(* IEC 61131-3 sources: moqui-plc/simatic-ax/src/moqui/framework/src/main/org/moqui/context, 9 files *)

(* ---- LogCmd.st ---- *)
TYPE LogCmd : (
    Idle, (* Waiting for commands *)
    Push (* Inserting a new log entry *)
); END_TYPE

(* ---- LogEvent.st ---- *)
TYPE LogEvent : STRUCT
	(* Unique identifier for the log event *)
    logEventId : STRING;
    loggerName : STRING;
	marker : LogMarker;
    level : LogLevel;
    logEventDate : DATE_AND_TIME;
	source : STRING;
	payloadType : LogPayloadType;
    payload : LogPayload;
	(* contextData: STRING; *)
	(*
	 * Occurrences this record stands for: 1 for an event, N for the summary that LoggerFacade writes when the
	 * same event was repeated N more times inside the suppression window ("last message repeated N times").
	 *)
    repeatCount : UINT;
	(* Position of the record in its LogRingBuffer, set by the buffer: consecutive records of one source differ by 1. *)
	sequence : UDINT;
END_STRUCT; END_TYPE

(* ---- LogLevel.st ---- *)
TYPE LogLevel : (
	Trace,
	Debug,
	Info,
	Warn,
	Error,
	Fatal,
	All,
	Off
); END_TYPE

(* ---- LogMarker.st ---- *)
TYPE LogMarker : (
	Diagnostics,
	Lifecycle,
	Integration,
	Health,
	Telemetry,
	AuditLog,
	Kpi,
	Measurement
); END_TYPE

(* ---- LogPayload.st ---- *)
TYPE LogPayload : STRUCT
	message : STRING;
    enumValue : UINT;
    numericValue : LREAL;
END_STRUCT; END_TYPE

(* ---- LogPayloadType.st ---- *)
TYPE LogPayloadType : (
    Text,
	Numeric,
	Enum
); END_TYPE

(* ---- LogSource.st ---- *)
(*
 * One registered LoggerFacade buffer, as seen by its consumer.
 * LoggerFacade sets logRef once; every other field belongs to the consumer. The AX port has no MQTT consumer yet
 * (the intended Siemens path is OPC UA): a future consumer follows LogDispatcher of the canonical IEC source.
 *)
TYPE LogSource : STRUCT
	(* Reference to log ring buffer *)
    logRef : REF_TO LogRingBuffer;
	(* Slot of the oldest record not yet released by the consumer *)
	readSlot : UINT := UINT#1;
	(* LogRingBuffer.droppedCount already reported by the consumer *)
	reportedDropCount : UDINT;
	(* Records published, and records discarded by the consumer *)
	publishedCount : UDINT;
	discardedCount : UDINT;
END_STRUCT; END_TYPE

(* ---- LoggerFacade.st ---- *)
USING System.Strings;

(*
 * Logger with local circular buffer and duplicate suppression.
 * Designed for central orchestration by a global LogAppender.
 *
 * - Level threshold: events below the global logMinLevel are ignored, as a log4j logger level.
 * - Duplicate suppression: an event equal to the last stored one (same logger, source, level, marker, payload
 *   type and value) within suppressDuration is only counted. The count is written later as one summary record,
 *   a copy of the event with repeatCount = repetitions, when a different event arrives or when the window has
 *   elapsed at any later call ("last message repeated N times"). Stored records are never modified.
 * - Rate limit: at most maxEventsPerWindow new events are stored in one suppressDuration window. Further
 *   events are only counted; at the first call after the window one Warn event reports how many were suppressed.
 *   Repetitions counted by duplicate suppression do not count against the limit.
 * - The local LogRingBuffer has this block as its only producer: call it from one task only.
 * - Inputs are retained between calls, as for every function block: pass level at every call,
 *   otherwise the event gets the level of the previous call.
 * - Generated logEventId: loggerName-<event sequence> (AX: no millisecond clock is read for the ID).
 *)
FUNCTION_BLOCK LoggerFacade
	VAR_EXTERNAL CONSTANT
		defaultLogLevel : LogLevel;
		defaultLogSuppressDuration : TIME;
		defaultLogSuppressDuplicates : BOOL;
		defaultLogMaxEventsPerWindow : UINT;
		LOG_SOURCE_LIST_MAX_SIZE : UINT;
	END_VAR
	VAR_EXTERNAL
		logSourceList : ARRAY[1..LOG_SOURCE_LIST_MAX_SIZE] OF LogSource;
		logSourceListSize : DINT;
		logMinLevel : LogLevel;
	END_VAR
	(* Log event data *)
	VAR_INPUT
		enable : BOOL;
		logEventId : STRING := '';
		loggerName : STRING;
		level : LogLevel := defaultLogLevel;
		marker : LogMarker := LogMarker#Diagnostics;
		source : STRING;
		payloadType : LogPayloadType := LogPayloadType#Text;
		message : STRING;
		enumValue : UINT;
		numericValue : LREAL;
	END_VAR
	(* Configuration parameters *)
	VAR_INPUT
		suppressDuplicates : BOOL := defaultLogSuppressDuplicates;
		suppressDuration : TIME := defaultLogSuppressDuration;
		(* Rate limit: new events stored per suppressDuration window (0 disables) *)
		maxEventsPerWindow : UINT := defaultLogMaxEventsPerWindow;
	END_VAR
	VAR_OUTPUT
		(* The event was stored, or counted as a repetition *)
		done : BOOL;
		(* The block could not register its buffer: LOG_SOURCE_LIST_MAX_SIZE is too small *)
		error : BOOL;
		(* The event, or a pending repetition summary, was refused because the local buffer was full *)
		dropped : BOOL;
		(* The event was not stored: the rate limit of the window was reached *)
		rateLimited : BOOL;
	END_VAR
	VAR
		(* Local log ring buffer *)
		logBuffer : LogRingBuffer;
		init : BOOL := FALSE;
		registered : BOOL;
		sourceSlot : DINT;
		isDuplicate : BOOL;
		now : DATE_AND_TIME;
		(* Last stored event, and repetitions of it not yet written *)
		lastLogEvent : LogEvent;
		hasLastLogEvent : BOOL;
		repeatPending : UINT;
		lastRepeatDate : DATE_AND_TIME;
		summary : LogEvent;
		eventRank : INT;
		minRank : INT;
		(* Log event ID generator *)
		eventSequence : UDINT := UDINT#0;
		(* Rate limit window *)
		windowOpen : BOOL;
		windowStart : DATE_AND_TIME;
		windowEventCount : UINT;
		windowSuppressed : UDINT;
		rateNotice : LogEvent;
	END_VAR

	done := FALSE;
	error := FALSE;
	dropped := FALSE;
	rateLimited := FALSE;

	(* Register once into the log appender source list *)
	IF NOT init THEN
		init := TRUE;
		logSourceListSize := logSourceListSize + DINT#1;
		sourceSlot := logSourceListSize;
		registered := (sourceSlot >= DINT#1) AND (sourceSlot <= TO_DINT(LOG_SOURCE_LIST_MAX_SIZE));
		IF registered THEN
			logSourceList[TO_UINT(sourceSlot)].logRef := REF(logBuffer);
		END_IF;
	END_IF;

	error := NOT registered;
	IF NOT enable OR NOT registered THEN RETURN; END_IF;

	now := nowTimestamp();

	(* Rate limit: at the end of the window report the suppressed events, then open a new window *)
	IF NOT windowOpen OR ((now - windowStart) >= suppressDuration) THEN
		IF (windowSuppressed > UDINT#0) AND (logMinLevel <> LogLevel#Off) THEN
			eventSequence := eventSequence + UDINT#1;
			rateNotice.logEventId := Concat(Concat(loggerName, '-suppressed-'), ToString(eventSequence));
			rateNotice.loggerName := loggerName;
			rateNotice.level := LogLevel#Warn;
			rateNotice.marker := LogMarker#Health;
			rateNotice.logEventDate := now;
			(* A device event, not a parameter value: empty source (DeviceLog of loggerName) *)
			rateNotice.source := '';
			rateNotice.payloadType := LogPayloadType#Text;
			rateNotice.payload.message := Concat(ToString(windowSuppressed), ' log events suppressed: logger too verbose');
			rateNotice.repeatCount := UINT#1;
			logBuffer(cmd := LogCmd#Push, logEntry := rateNotice);
			logBuffer.cmd := LogCmd#Idle;
			dropped := logBuffer.dropped;
		END_IF;
		windowOpen := TRUE;
		windowStart := now;
		windowEventCount := UINT#0;
		windowSuppressed := UDINT#0;
	END_IF;

	(* Write the pending repetition summary once its window has elapsed *)
	IF (repeatPending > UINT#0) AND ((now - lastLogEvent.logEventDate) >= suppressDuration) THEN
		summary := lastLogEvent;
		summary.logEventId := Concat(lastLogEvent.logEventId, '-repeated');
		summary.logEventDate := lastRepeatDate;
		summary.repeatCount := repeatPending;
		repeatPending := UINT#0;
		logBuffer(cmd := LogCmd#Push, logEntry := summary);
		dropped := dropped OR logBuffer.dropped;
	END_IF;

	(* Level threshold: All is the lowest threshold, Off disables logging *)
	CASE level OF
		LogLevel#Trace: eventRank := INT#0;
		LogLevel#Debug: eventRank := INT#1;
		LogLevel#Info: eventRank := INT#2;
		LogLevel#Warn: eventRank := INT#3;
		LogLevel#Error: eventRank := INT#4;
		LogLevel#Fatal: eventRank := INT#5;
	ELSE
		eventRank := INT#-1;
	END_CASE;
	CASE logMinLevel OF
		LogLevel#Trace, LogLevel#All: minRank := INT#0;
		LogLevel#Debug: minRank := INT#1;
		LogLevel#Info: minRank := INT#2;
		LogLevel#Warn: minRank := INT#3;
		LogLevel#Error: minRank := INT#4;
		LogLevel#Fatal: minRank := INT#5;
	ELSE
		minRank := INT#6;
	END_CASE;
	IF (eventRank < INT#0) OR (eventRank < minRank) THEN RETURN; END_IF;

	(* Compression logic (duplicate suppression) *)
	isDuplicate := FALSE;
	IF hasLastLogEvent AND suppressDuplicates AND (payloadType = lastLogEvent.payloadType)
			AND (loggerName = lastLogEvent.loggerName)
			AND (source = lastLogEvent.source)
			AND (level = lastLogEvent.level)
			AND (marker = lastLogEvent.marker)
			AND ((now - lastLogEvent.logEventDate) < suppressDuration) THEN
		CASE payloadType OF
			LogPayloadType#Text: isDuplicate := (message = lastLogEvent.payload.message);
			LogPayloadType#Enum: isDuplicate := (enumValue = lastLogEvent.payload.enumValue);
			LogPayloadType#Numeric: isDuplicate := (numericValue = lastLogEvent.payload.numericValue);
		END_CASE;
	END_IF;

	IF isDuplicate THEN
		(* Count the repetition; the summary record is written later *)
		IF repeatPending < UINT#65535 THEN repeatPending := repeatPending + UINT#1; END_IF;
		lastRepeatDate := now;
		done := TRUE;
		RETURN;
	END_IF;

	(*
	 * Rate limit: over the limit the new event is only counted. Checked before the repetition summary,
	 * so alternating events cannot write one summary per call; the summary is written when the window elapses.
	 *)
	IF (maxEventsPerWindow > UINT#0) AND (windowEventCount >= maxEventsPerWindow) THEN
		IF windowSuppressed < UDINT#16#FFFFFFFF THEN windowSuppressed := windowSuppressed + UDINT#1; END_IF;
		rateLimited := TRUE;
		RETURN;
	END_IF;
	windowEventCount := windowEventCount + UINT#1;

	(* A different event: first write the repetitions of the previous one *)
	IF repeatPending > UINT#0 THEN
		summary := lastLogEvent;
		summary.logEventId := Concat(lastLogEvent.logEventId, '-repeated');
		summary.logEventDate := lastRepeatDate;
		summary.repeatCount := repeatPending;
		repeatPending := UINT#0;
		logBuffer(cmd := LogCmd#Push, logEntry := summary);
		dropped := dropped OR logBuffer.dropped;
	END_IF;

	(* Prepare the new log event entry *)
	IF logEventId = '' THEN
		eventSequence := eventSequence + UDINT#1;
		lastLogEvent.logEventId := Concat(Concat(loggerName, '-'), ToString(eventSequence));
	ELSE
		lastLogEvent.logEventId := logEventId;
	END_IF;

	lastLogEvent.loggerName := loggerName;
	lastLogEvent.level := level;
	lastLogEvent.marker := marker;
	lastLogEvent.logEventDate := now;
	lastLogEvent.source := source;
	lastLogEvent.payloadType := payloadType;
	lastLogEvent.repeatCount := UINT#1;

	CASE payloadType OF
		LogPayloadType#Text: lastLogEvent.payload.message := message;
		LogPayloadType#Enum: lastLogEvent.payload.enumValue := enumValue;
		LogPayloadType#Numeric: lastLogEvent.payload.numericValue := numericValue;
	END_CASE;

	(* Append the new log event *)
	logBuffer(cmd := LogCmd#Push, logEntry := lastLogEvent);
	logBuffer.cmd := LogCmd#Idle;

	done := logBuffer.done;
	dropped := dropped OR logBuffer.dropped;
	(* A refused event must not be followed by repetitions of it: the next equal event is stored as new *)
	hasLastLogEvent := logBuffer.done;
END_FUNCTION_BLOCK

(* ---- LogRingBuffer.st ---- *)
(*
 * Bounded log queue between one producer and one consumer, without locks and without waits.
 *
 * - Producer: the LoggerFacade that owns this instance, in its own task. It calls the block with cmd := LogCmd#Push,
 *   writes logBuffer[writeSlot] and only then publishes the record by incrementing writeCount.
 * - Consumer: reads the records between readCount and writeCount, starting from its LogSource.readSlot, and
 *   releases them by incrementing readCount. The AX port has no consumer yet: the queue fills and then refuses.
 *
 * Each counter has a single writer. The S7-1500 runs the user program on one core and a 32-bit aligned write is
 * atomic, so a task that preempts another sees the counters in program order; the canonical CODESYS source uses
 * __XADD for multicore targets. When the queue is full the new record is refused and counted in droppedCount.
 *)
FUNCTION_BLOCK LogRingBuffer
	VAR_EXTERNAL CONSTANT
	    LOG_MAX_SIZE : UINT;
	END_VAR
	VAR_INPUT
	    cmd : LogCmd := LogCmd#Idle;
	    logEntry : LogEvent;
	END_VAR
	VAR_OUTPUT
	    done : BOOL;
	    error : BOOL;
	    (* The record was refused because the queue was full *)
	    dropped : BOOL;
	    logBuffer : ARRAY[1..LOG_MAX_SIZE] OF LogEvent;
	    (* Records ever written (producer-owned); wraps around, only differences are meaningful *)
	    writeCount : DINT;
	    (* Records ever released (consumer-owned) *)
	    readCount : DINT;
	    (* Records refused because the queue was full (producer-owned) *)
	    droppedCount : UDINT;
	    isFull : BOOL;
	    isEmpty : BOOL;
	END_VAR
	VAR
	    writeSlot : UINT := UINT#1;
	    pending : DINT;
	END_VAR

	done := FALSE;
	error := FALSE;
	dropped := FALSE;

	IF cmd = LogCmd#Idle THEN RETURN; END_IF;
	IF (cmd <> LogCmd#Push) OR (writeSlot < UINT#1) OR (writeSlot > LOG_MAX_SIZE) THEN
	    error := TRUE;
	    RETURN;
	END_IF;

	pending := writeCount - readCount;
	IF (pending < DINT#0) OR (pending >= TO_DINT(LOG_MAX_SIZE)) THEN
	    (* Full, or counters out of range: refuse the record, never overwrite unreleased records *)
	    IF droppedCount < UDINT#16#FFFFFFFF THEN droppedCount := droppedCount + UDINT#1; END_IF;
	    dropped := TRUE;
	    isFull := TRUE;
	    isEmpty := FALSE;
	    RETURN;
	END_IF;

	logBuffer[writeSlot] := logEntry;
	logBuffer[writeSlot].sequence := TO_UDINT(writeCount) + UDINT#1;
	writeSlot := (writeSlot MOD LOG_MAX_SIZE) + UINT#1;
	(* Publish the record after it is complete *)
	writeCount := writeCount + DINT#1;
	done := TRUE;

	isFull := (pending + DINT#1) >= TO_DINT(LOG_MAX_SIZE);
	isEmpty := FALSE;
END_FUNCTION_BLOCK
